{attribute 'no_assign'}
FUNCTION_BLOCK FB_DO_WTURBINE_LD0_WTUR1_DmdWSpt EXTENDS FB_AcsiCommonDataClass
VAR_INPUT
	val: FB_DO_WTURBINE_LD0_WTUR1_DmdWSpt_val := (sClass:='APC', bLinkResult:=THIS^.AddDataToContainer(ipData:=val));
END_VAR
VAR
END_VAR

END_FUNCTION_BLOCK

(* stored: Version 1.1.0.1
   POU FB_DO_WTURBINE_LD0_WTUR1_DmdWSpt: Id {c3faf58c-cd53-43c7-841f-9b14c56404a4}, SpecialFunc None *)
